Fanuc KAREL source: kc00045.KL

-- PROVISIONAL review KL for V1013-1; original PC SHA256 1d52ada140572cd72cf818a7ed19e82cc0dd3c2d7b0911cb1b262cc79b1bfd69
-- Incomplete behavior may be omitted. Consult companion uncertainty JSON. Do not deploy.
PROGRAM KC00045
%NOLOCKGROUP
BEGIN
  -- UNRESOLVED_PC offsets 5-29; opcodes 27,22,22,2A,22,31
  -- UNRESOLVED_PC offsets 34-38; opcodes 7F
END KC00045
